TYPE ST_Axis :
STRUCT
    fPos : LREAL;
    fVel : LREAL;
END_STRUCT
END_TYPE

(* stored: Version 1.1.0.1, ProductVersion 3.1.4024.12
   DUT ST_Axis: Id {bbbbbbbb-0000-0000-0000-000000000001} *)
